// TwinCAT 3 PLC project PlcSafety
// ProgramVersion: 3.1.4026.27
// CompilerDefines: VISU_USEPROPERTYINFO
// libraries:
//   Tc2_Standard, * (Beckhoff Automation GmbH)
//   Tc2_System, * (Beckhoff Automation GmbH)
//   VisuDialogs, * (System)
// project tree:
//   / GlobalTextList.TcGTLO, PlcTask.TcTTO, Visualization Manager.TcVMO (not stored)
//   GVLs/ GVL_Safety.TcGVL
//   POUs/ MAIN.TcPOU, PRG_SafetyInterface.TcPOU
//   VISUs/ VISU_SafetySim.TcVIS
// real-time tasks:
//   TASK PlcTask: cycle T#10ms, priority 20, ADS port 350
// I/O:
//   DEVICE Device 1 (EtherCAT) (disabled), AmsNetId 192.168.1.24.2.1
//     Term 1 (EK1100) [EK1100 EtherCAT Coupler (2A E-Bus)]
//       Term 2 (EL6910) [EL6910, TwinSAFE PLC]
//       Term 3 (EL1904) [EL1904, 4 Ch. Safety Input 24V, TwinSAFE]
//         modules: Module 1 (FSOES)
//       Term 4 (EL2904) [EL2904, 4 Ch. Safety Output 24V, 0.5A, TwinSAFE]
//         modules: Module 1 (FSOES), Module 2 (DO)
// variable links:
//   (this object) <-> Device 1 (EtherCAT)
//     Term 1 (EK1100)/Term 2 (EL6910)/ConnectionInputs/TwinSafeGroup1.EStop1_In_3 TxPDO <-> Term 1 (EK1100)/Term 3 (EL1904)/Module 1 (FSOES)/RxPDO/FSOE
//     Term 1 (EK1100)/Term 2 (EL6910)/ConnectionInputs/TwinSafeGroup1.EStop1_Out_4 TxPDO <-> Term 1 (EK1100)/Term 4 (EL2904)/Module 1 (FSOES)/RxPDO/FSOE
//     Term 1 (EK1100)/Term 2 (EL6910)/ConnectionOutputs/TwinSafeGroup1.EStop1_In_3 RxPDO <-> Term 1 (EK1100)/Term 3 (EL1904)/Module 1 (FSOES)/TxPDO/FSOE
//     Term 1 (EK1100)/Term 2 (EL6910)/ConnectionOutputs/TwinSafeGroup1.EStop1_Out_4 RxPDO <-> Term 1 (EK1100)/Term 4 (EL2904)/Module 1 (FSOES)/TxPDO/FSOE
//     Term 1 (EK1100)/Term 3 (EL1904)/Module 1 (FSOES)/RxPDO/FSOE <-> Term 1 (EK1100)/Term 2 (EL6910)/ConnectionInputs/TwinSafeGroup1.EStop1_In_3 TxPDO
//     Term 1 (EK1100)/Term 3 (EL1904)/Module 1 (FSOES)/TxPDO/FSOE <-> Term 1 (EK1100)/Term 2 (EL6910)/ConnectionOutputs/TwinSafeGroup1.EStop1_In_3 RxPDO
//     Term 1 (EK1100)/Term 4 (EL2904)/Module 1 (FSOES)/RxPDO/FSOE <-> Term 1 (EK1100)/Term 2 (EL6910)/ConnectionInputs/TwinSafeGroup1.EStop1_Out_4 TxPDO
//     Term 1 (EK1100)/Term 4 (EL2904)/Module 1 (FSOES)/TxPDO/FSOE <-> Term 1 (EK1100)/Term 2 (EL6910)/ConnectionOutputs/TwinSafeGroup1.EStop1_Out_4 RxPDO
//   (this object) <-> Device 1 (EtherCAT)/Term 1 (EK1100)/Term 2 (EL6910)
//     PlcTask Inputs/GVL_Safety.bEStop1_SafeHealthy <-> StandardInputs/TwinSafeGroup1.EStop1_SafeHealthy_6
//     PlcTask Inputs/GVL_Safety.bSafety_ComFault <-> StandardInputs/TwinSafeGroup1.Safety_ComFault_7
//     PlcTask Outputs/GVL_Safety.bEStop1_RestartOut <-> StandardOutputs/TwinSafeGroup1.EStop1_Restart_5
//     PlcTask Outputs/GVL_Safety.bSafety_ErrAckOut <-> StandardOutputs/TwinSafeGroup1.ErrorAcknowledgement_1
//     PlcTask Outputs/GVL_Safety.bSafety_GroupRunOut <-> StandardOutputs/TwinSafeGroup1.Run_2

CONFIGURATION PlcSafety
    RESOURCE PLC ON TwinCAT3
        TASK PlcTask(INTERVAL := T#10ms, PRIORITY := 20);
        PROGRAM MAIN WITH PlcTask : MAIN;
    END_RESOURCE
END_CONFIGURATION

// ---- GVLs/GVL_Safety.TcGVL
{attribute 'qualified_only'}
VAR_GLOBAL
    // Operator / HMI / sequence commands (internal PLC tags)
    bEStop1_ResetCmd     : BOOL;         // Momentary reset request from HMI/button
    bSafety_ErrAckCmd    : BOOL;         // Momentary error acknowledge request

    // Rising-edge outputs mapped to TwinSAFE standard aliases (PLC -> TwinSAFE)
    bEStop1_RestartOut   AT %Q* : BOOL;  // Linked to EStop1_Restart.sds
    bSafety_ErrAckOut    AT %Q* : BOOL;  // Linked to ErrorAcknowledgement.sds
    bSafety_GroupRunOut  AT %Q* : BOOL;  // Linked to Run.sds (TwinSAFE group run enable)

    // Safety status & diagnostics (TwinSAFE / I/O -> PLC)
    bEStop1_SafeHealthy  AT %I* : BOOL;  // TRUE when E-Stop safe output is healthy
    bEStop1_Tripped      : BOOL;         // Derived: TRUE when E-Stop is open/tripped
    bSafety_ComFault     AT %I* : BOOL;  // Safety communication / group fault status
END_VAR

// ---- POUs/MAIN.TcPOU
PROGRAM MAIN
VAR
END_VAR

PRG_SafetyInterface();

END_PROGRAM

// ---- POUs/PRG_SafetyInterface.TcPOU
PROGRAM PRG_SafetyInterface
VAR
    fbResetPulse  : R_TRIG;
    fbErrAckPulse : R_TRIG;
END_VAR

// Single-scan rising-edge pulse so Restart never stays stuck TRUE
fbResetPulse(CLK := GVL_Safety.bEStop1_ResetCmd);
GVL_Safety.bEStop1_RestartOut := fbResetPulse.Q;

// Single-scan rising-edge pulse for TwinSAFE group error acknowledgment
fbErrAckPulse(CLK := GVL_Safety.bSafety_ErrAckCmd);
GVL_Safety.bSafety_ErrAckOut := fbErrAckPulse.Q;

// Derive machine-side tripped state from safe output status
GVL_Safety.bEStop1_Tripped := NOT GVL_Safety.bEStop1_SafeHealthy;

// Keep TwinSAFE group run signal enabled during normal PLC execution
GVL_Safety.bSafety_GroupRunOut := TRUE;

END_PROGRAM

// ---- GlobalTextList.TcGTLO
TEXTLIST GlobalTextList
  497 = 'Ack Fault'
  635 = 'Commands'
  394 = 'ErrAckOut (Pulse)'
  7 = 'EStop1 SafeHealthy'
  756 = 'EStop1 Tripped'
  993 = 'Reset E-Stop'
  670 = 'RestartOut (Pulse)'
  863 = 'Safety ComFault'
  777 = 'Status'
END_TEXTLIST

// ---- VISUs/VISU_SafetySim.TcVIS
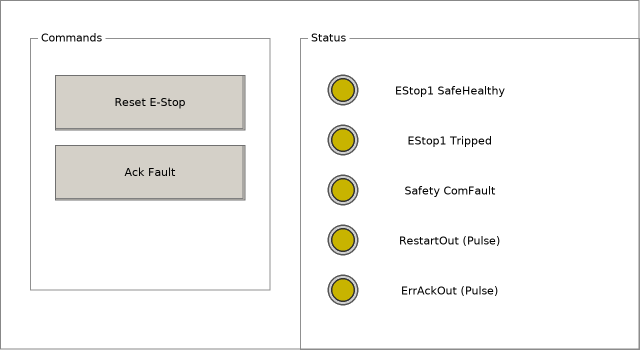
VISUALIZATION VISU_SafetySim  // 640x350
    GroupBox (300,30 340x320), "Status"
    GroupBox (30,30 240x260), "Commands"
    Lamp1 (325,72 36x36), variable: GVL_Safety.bEStop1_SafeHealthy, style: Lamp-Lamp1-Yellow
    Label (375,76 150x30), "EStop1 SafeHealthy"
    Label (375,176 150x30), "Safety ComFault"
    Label (375,126 150x30), "EStop1 Tripped"
    Label (375,276 150x30), "ErrAckOut (Pulse)"
    Label (375,226 150x30), "RestartOut (Pulse)"
    Lamp1 (325,122 36x36), variable: GVL_Safety.bEStop1_Tripped, style: Lamp-Lamp1-Yellow
    Lamp1 (325,172 36x36), variable: GVL_Safety.bSafety_ComFault, style: Lamp-Lamp1-Yellow
    Lamp1 (325,272 36x36), variable: GVL_Safety.bSafety_ErrAckOut, style: Lamp-Lamp1-Yellow
    Lamp1 (325,222 36x36), variable: GVL_Safety.bEStop1_RestartOut, style: Lamp-Lamp1-Yellow
    Button (55,75 190x55), "Reset E-Stop", pressed state: GVL_Safety.bEStop1_ResetCmd
        tap GVL_Safety.bEStop1_ResetCmd
    Button (55,145 190x55), "Ack Fault", pressed state: GVL_Safety.bSafety_ErrAckCmd
        tap GVL_Safety.bSafety_ErrAckCmd
END_VISUALIZATION
